(* IEC 61131-3 sources: sis-interlock-demo/tests/POUs/Suites/FB_SisUtil_Test, 5 files *)

(* ---- CemCrcDemoMatrixValue.method.decl.st ---- *)
// CRC матрицы демо-объекта (10 причин, 7 следствий, маски таблицы 11.4) — 16#CD40; локальная копия
// масок, а не GVL_SisCfg: тест не зависит от сгенерированного кода
METHOD PRIVATE CemCrcDemoMatrixValue
VAR
    stCfg : ST_CemCfg;   // матрица демо-объекта (только счётчики и маски)
END_VAR

(* ---- Crc16CheckValue.method.decl.st ---- *)
// Контрольное значение CRC-16/CCITT-FALSE: ASCII «123456789» → 16#29B1
METHOD PRIVATE Crc16CheckValue
VAR
    wCrc : WORD;    // регистр CRC
    uiCh : UINT;    // код очередного символа
END_VAR

(* ---- Crc16CheckValue.method.impl.st ---- *)
coUnit.TEST('Sis_Crc16_CheckValue');
wCrc := GVL_Const.CRC16_INIT;
FOR uiCh := 16#31 TO 16#39 DO
    wCrc := F_SisCrc16Byte(wCrc := wCrc, bData := UINT_TO_BYTE(uiCh));
END_FOR
AssertEquals_WORD(Expected := 16#29B1, Actual := wCrc, Message := 'CRC-16/CCITT-FALSE of 123456789');
coUnit.TEST_FINISHED();

(* ---- LogEventNoSinkReturnsFalse.method.decl.st ---- *)
// F_SisLogEvent: без приёмника — FALSE; с приёмником — TRUE, поля записи переданы, номер — от журнала
METHOD PRIVATE LogEventNoSinkReturnsFalse
VAR
    fbLog   : FB_SisEventLog;   // журнал
    itfNone : I_SisEventSink;   // пустая ссылка
    xRes    : BOOL;             // результат
    stEv    : ST_SisEvent;      // последнее событие
END_VAR

(* ---- Ne43ValidLimits.method.decl.st ---- *)
// F_SisNe43Valid: 3,6 и 21,0 мА — недостоверно, 3,61 и 20,99 мА — достоверно, NaN и 0 мА — нет
METHOD PRIVATE Ne43ValidLimits
VAR
    uBits : PL.U_RealBits;   // значение REAL по битам IEEE 754
END_VAR
